Fanuc KAREL source: KO00076.KL

PROGRAM KO00076
%NOLOCKGROUP
%ENVIRONMENT MIR
VAR
  P1: XYZWPREXT
  P2: XYZWPREXT
  F: BOOLEAN
  OUT: JOINTPOS
BEGIN
  F = TRUE
  OUT = MIRROR(P1, P2, F)
END KO00076
